Omron Sysmac Studio project ENG3106C Project (Sysmac Studio 1.60.0.64010, StandardProject)
(* This is the project *)

# Controller PLC0: NX102-1020 version 1.48
Units and slaves: Unit 1 : NX-PF0630 (N1); Unit 2 : NX-ID5142-1 (N2); Unit 3 : NX-OC4633 (N3)
Task PrimaryTask (priority 4, period or condition 2000): Main

TYPE sql_equipment : STRUCT
    equip_id : STRING[128];
    equip_name : STRING[128];
    current_equip_state : STRING[128];
    former_equip_state : STRING[128];
    former_lot_id : STRING[128];
    upd_dt : DATE_AND_TIME;
    current_station_id : STRING[128];
END_STRUCT END_TYPE
TYPE sql_event_history : STRUCT
    event_id : STRING[128];
    request_id : STRING[128];
    equip_id : STRING[128];
    start_dt : DATE_AND_TIME;
    end_dt : DATE_AND_TIME;
    source_location : STRING[128];
    destination_location : STRING[128];
    request_client : STRING[128];
    event_type : STRING[128];
    time_taken_seconds : INT;
END_STRUCT END_TYPE
TYPE sql_lot : STRUCT
    lot_id : STRING[128];
    product_name : STRING[128];
    lot_status : STRING[128];
    create_dt : DATE_AND_TIME;
END_STRUCT END_TYPE
TYPE sql_request_details : STRUCT
    request_id : STRING[128];
    operating_start_dt : DATE_AND_TIME;
    operating_end_dt : DATE_AND_TIME;
    equip_id : STRING[128];
    target_location : STRING[128];
    home_location : STRING[128];
    request_state : STRING[128];
END_STRUCT END_TYPE
TYPE sql_station : STRUCT
    station_id : STRING[128];
    station_name : STRING[128];
    station_type : STRING[128];
END_STRUCT END_TYPE

VAR_GLOBAL
    gInput01 : BOOL;  (* at IOBus://unit#2/Input Bit 16 bits/Input Bit 01 *)
    gInput00 : BOOL;  (* at IOBus://unit#2/Input Bit 16 bits/Input Bit 00 *)
    gInput02 : BOOL;  (* at IOBus://unit#2/Input Bit 16 bits/Input Bit 02 *)
    gInput06 : BOOL;  (* at IOBus://unit#2/Input Bit 16 bits/Input Bit 06 *)
    gInput07 : BOOL;  (* at IOBus://unit#2/Input Bit 16 bits/Input Bit 07 *)
    gInput08 : BOOL;  (* at IOBus://unit#2/Input Bit 16 bits/Input Bit 08 *)
    gInput09 : BOOL;  (* at IOBus://unit#2/Input Bit 16 bits/Input Bit 09 *)
    gInput10 : BOOL;  (* at IOBus://unit#2/Input Bit 16 bits/Input Bit 10 *)
    gInput11 : BOOL;  (* at IOBus://unit#2/Input Bit 16 bits/Input Bit 11 *)
    gPB13 : BOOL;  (* at IOBus://unit#2/Input Bit 16 bits/Input Bit 13 *)
    gPB14 : BOOL;  (* at IOBus://unit#2/Input Bit 16 bits/Input Bit 14 *)
    gPB15 : BOOL;  (* at IOBus://unit#2/Input Bit 16 bits/Input Bit 15 *)
    gOutput00 : BOOL;  (* at IOBus://unit#3/Output Bit 8 bits/Output Bit 00 *)
    gOutput01 : BOOL;  (* at IOBus://unit#3/Output Bit 8 bits/Output Bit 01 *)
    gOutput02 : BOOL;  (* at IOBus://unit#3/Output Bit 8 bits/Output Bit 02 *)
    gOutput03 : BOOL;  (* at IOBus://unit#3/Output Bit 8 bits/Output Bit 03 *)
    gOutput04 : BOOL;  (* at IOBus://unit#3/Output Bit 8 bits/Output Bit 04 *)
    gOutput05 : BOOL;  (* at IOBus://unit#3/Output Bit 8 bits/Output Bit 05 *)
    gOutput06 : BOOL;  (* at IOBus://unit#3/Output Bit 8 bits/Output Bit 06 *)
    gOutput07 : BOOL;  (* at IOBus://unit#3/Output Bit 8 bits/Output Bit 07 *)
    gStart : BOOL;
    gStop : BOOL;
    gMachineOn : BOOL;
    gStartB : BOOL;  (* published *)
    gStartA : BOOL;  (* published *)
    gGoOutBase : BOOL;  (* published *)
    gGoBackBase : BOOL;  (* published *)
    gSessionTransferSuccess : INT;  (* published *)
    gSessionMotorUsageElapsed : INT;  (* published *)
    gProgressA : BOOL;
    gProgressB : BOOL;
END_VAR

PROGRAM Main
VAR
    Step4 : RS;
    gMotorClockwise : BOOL;
    gMotorCounterClockwise : BOOL;
    Step5 : RS;
    Step6 : RS;
    StationA : RS;
    StationB : RS;
    DB_Connect_instance : DB_Connect;
    AmhsDb1 : DWORD;
    test1 : BOOL;
    test2 : BOOL;
    DB_CreateMapping_instance : DB_CreateMapping;
    test3 : BOOL;
    DB_Close_instance : DB_Close;
    Step1B : RS;
    Step1A : RS;
    Step2A : RS;
    Step2B : RS;
    Step3A : RS;
    Step3B : RS;
    Timer1A : TON;
    Timer1B : TON;
    Timer4 : TON;
    DB_Insert_instance : DB_Insert;
    test_map_varr : sql_event_history;
    test4 : BOOL;
    test5 : BOOL;
    Step0A : RS;
    Step0B : RS;
    Counter1 : CTU;
END_VAR
VAR_EXTERNAL
    gPB13 : BOOL;
    gPB14 : BOOL;
    gMachineOn : BOOL;
    gOutput06 : BOOL;
    gOutput07 : BOOL;
    gInput01 : BOOL;
    gOutput00 : BOOL;
    gOutput01 : BOOL;
    gOutput04 : BOOL;
    gOutput05 : BOOL;
    gInput07 : BOOL;
    gInput06 : BOOL;
    gInput00 : BOOL;
    gInput11 : BOOL;
    gInput10 : BOOL;
    gStartA : BOOL;
    gStartB : BOOL;
    gInput02 : BOOL;
    gInput09 : BOOL;
    gInput08 : BOOL;
    gOutput02 : BOOL;
    gOutput03 : BOOL;
    gGoOutBase : BOOL;
    gGoBackBase : BOOL;
    gPB15 : BOOL;
    gProgressA : BOOL;
    gProgressB : BOOL;
END_VAR
VAR
    _e1 : R_TRIG;
    _e2 : R_TRIG;
    _e3 : F_TRIG;
    _e4 : F_TRIG;
    _e5 : F_TRIG;
    _e6 : F_TRIG;
    _e7 : F_TRIG;
    _e8 : F_TRIG;
    _e9 : F_TRIG;
    _e10 : F_TRIG;
    _p11 : BOOL;
    _e12 : R_TRIG;
END_VAR

(* Section Section0: ladder, written here as Structured Text *)

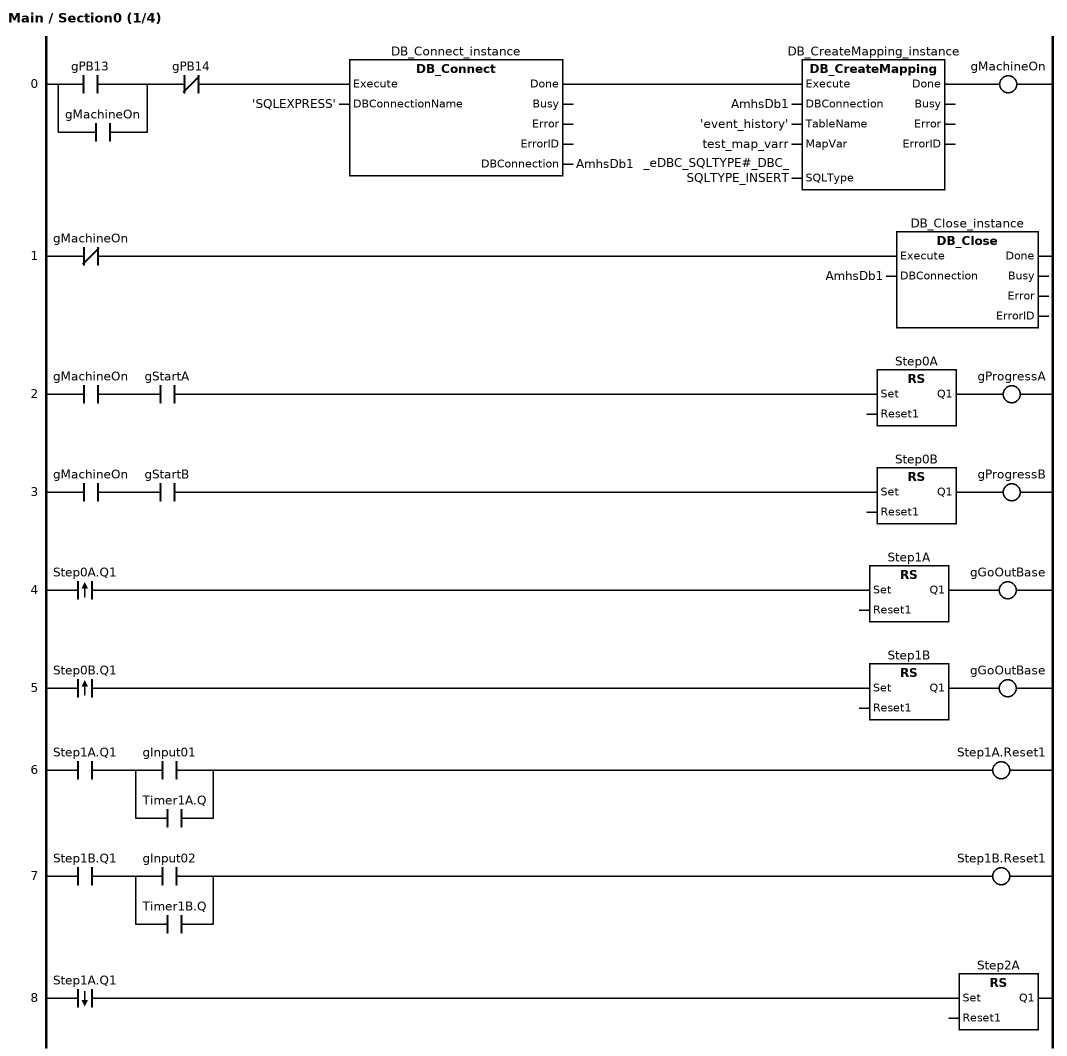
(* Rung 0 *)
DB_Connect_instance(Execute := (gPB13 OR gMachineOn) AND NOT gPB14, DBConnectionName := 'SQLEXPRESS', DBConnection => AmhsDb1);
DB_CreateMapping_instance(Execute := DB_Connect_instance.Done, DBConnection := AmhsDb1, TableName := 'event_history', MapVar := test_map_varr, SQLType := _eDBC_SQLTYPE#_DBC_SQLTYPE_INSERT);
gMachineOn := DB_CreateMapping_instance.Done;
(* Rung 1 *)
DB_Close_instance(Execute := NOT gMachineOn, DBConnection := AmhsDb1);
(* Rung 2 *)
Step0A(Set := gMachineOn AND gStartA);
gProgressA := Step0A.Q1;
(* Rung 3 *)
Step0B(Set := gMachineOn AND gStartB);
gProgressB := Step0B.Q1;
(* Rung 4 *)
_e1(CLK := Step0A.Q1);
Step1A(Set := _e1.Q);
gGoOutBase := Step1A.Q1;
(* Rung 5 *)
_e2(CLK := Step0B.Q1);
Step1B(Set := _e2.Q);
gGoOutBase := Step1B.Q1;
(* Rung 6 *)
Step1A.Reset1 := Step1A.Q1 AND (gInput01 OR Timer1A.Q);
(* Rung 7 *)
Step1B.Reset1 := Step1B.Q1 AND (gInput02 OR Timer1B.Q);
(* Rung 8 *)
_e3(CLK := Step1A.Q1);
Step2A(Set := _e3.Q);

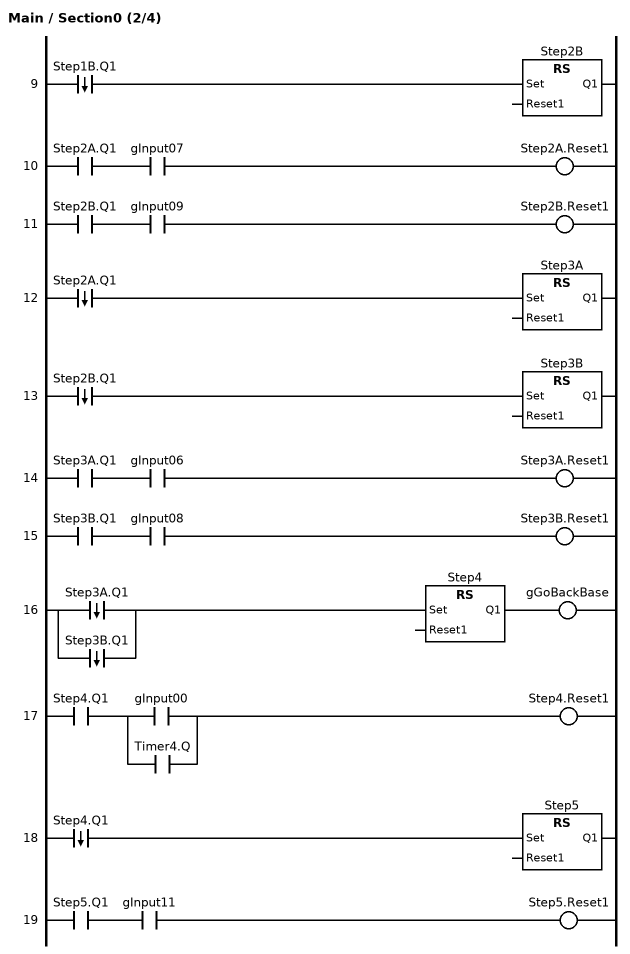
(* Rung 9 *)
_e4(CLK := Step1B.Q1);
Step2B(Set := _e4.Q);
(* Rung 10 *)
Step2A.Reset1 := Step2A.Q1 AND gInput07;
(* Rung 11 *)
Step2B.Reset1 := Step2B.Q1 AND gInput09;
(* Rung 12 *)
_e5(CLK := Step2A.Q1);
Step3A(Set := _e5.Q);
(* Rung 13 *)
_e6(CLK := Step2B.Q1);
Step3B(Set := _e6.Q);
(* Rung 14 *)
Step3A.Reset1 := Step3A.Q1 AND gInput06;
(* Rung 15 *)
Step3B.Reset1 := Step3B.Q1 AND gInput08;
(* Rung 16 *)
_e7(CLK := Step3A.Q1);
_e8(CLK := Step3B.Q1);
Step4(Set := _e7.Q OR _e8.Q);
gGoBackBase := Step4.Q1;
(* Rung 17 *)
Step4.Reset1 := Step4.Q1 AND (gInput00 OR Timer4.Q);
(* Rung 18 *)
_e9(CLK := Step4.Q1);
Step5(Set := _e9.Q);
(* Rung 19 *)
Step5.Reset1 := Step5.Q1 AND gInput11;

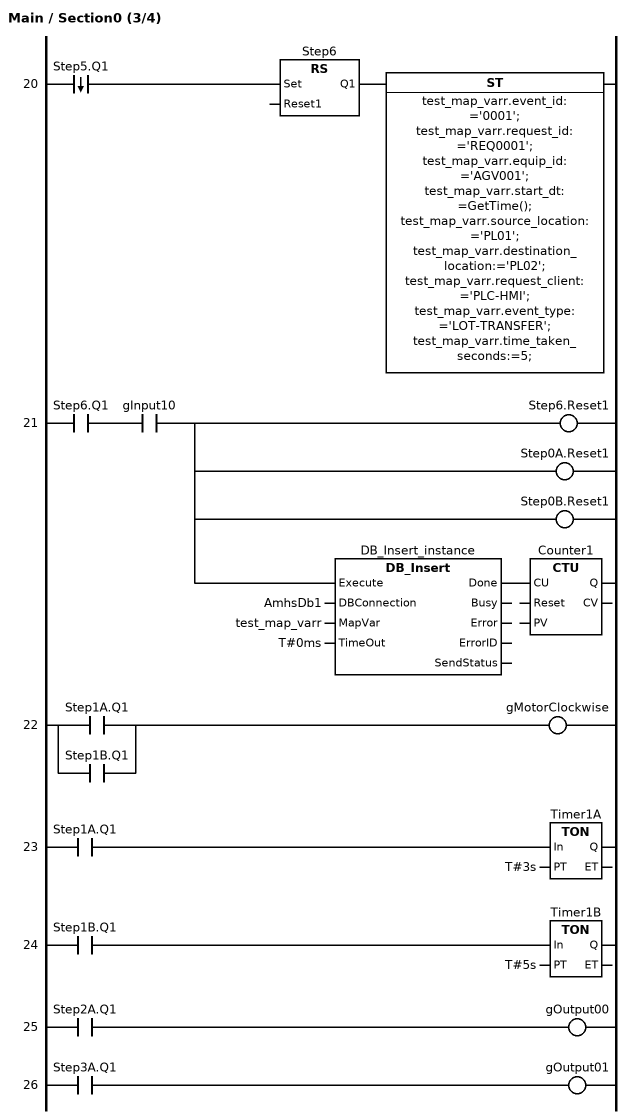
(* Rung 20 *)
_e10(CLK := Step5.Q1);
Step6(Set := _e10.Q);
IF Step6.Q1 THEN
    test_map_varr.event_id:='0001';
    test_map_varr.request_id:='REQ0001';
    test_map_varr.equip_id:='AGV001';
    test_map_varr.start_dt:=GetTime();
    test_map_varr.source_location:='PL01';
    test_map_varr.destination_location:='PL02';
    test_map_varr.request_client:='PLC-HMI';
    test_map_varr.event_type:='LOT-TRANSFER';
    test_map_varr.time_taken_seconds:=5;
END_IF;
(* Rung 21 *)
_p11 := Step6.Q1 AND gInput10;
Step6.Reset1 := _p11;
Step0A.Reset1 := _p11;
Step0B.Reset1 := _p11;
DB_Insert_instance(Execute := _p11, DBConnection := AmhsDb1, MapVar := test_map_varr, TimeOut := T#0ms);
_e12(CLK := DB_Insert_instance.Done);
Counter1(CU := _e12.Q);
(* Rung 22 *)
gMotorClockwise := Step1A.Q1 OR Step1B.Q1;
(* Rung 23 *)
Timer1A(In := Step1A.Q1, PT := T#3s);
(* Rung 24 *)
Timer1B(In := Step1B.Q1, PT := T#5s);
(* Rung 25 *)
gOutput00 := Step2A.Q1;
(* Rung 26 *)
gOutput01 := Step3A.Q1;

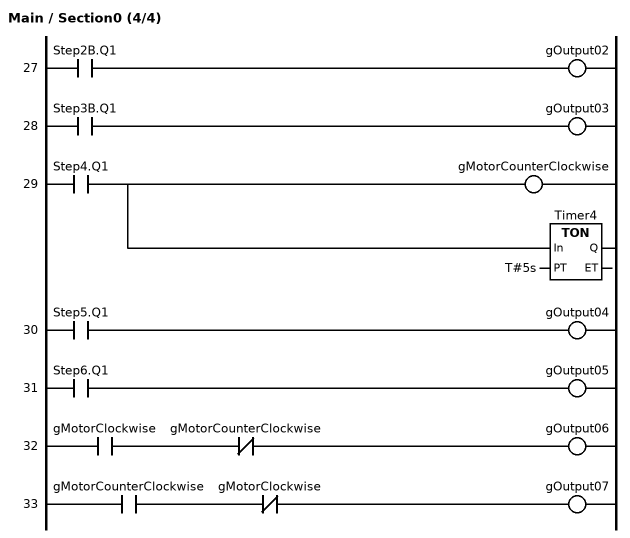
(* Rung 27 *)
gOutput02 := Step2B.Q1;
(* Rung 28 *)
gOutput03 := Step3B.Q1;
(* Rung 29 *)
gMotorCounterClockwise := Step4.Q1;
Timer4(In := Step4.Q1, PT := T#5s);
(* Rung 30 *)
gOutput04 := Step5.Q1;
(* Rung 31 *)
gOutput05 := Step6.Q1;
(* Rung 32 *)
gOutput06 := gMotorClockwise AND NOT gMotorCounterClockwise;
(* Rung 33 *)
gOutput07 := gMotorCounterClockwise AND NOT gMotorClockwise;
END_PROGRAM

# Device HMI_NA5_0 (NA): not converted